// TIA Portal V20 export
// export: Created 2026-10-19T18:45:22.4932904Z, ExportSetting None, DisplayName Totally Integrated Automation Portal, DisplayVersion V20 Update 6, DisplayName TIA Portal Openness, DisplayVersion V20 Update 6, DisplayName TIA Portal Version Control Interface, DisplayVersion V20 Update 6, DisplayName SINAMICS Startdrive Advanced, DisplayVersion V20 SP1, DisplayName SINAMICS Startdrive G130, G150, S120, S150, SINAMICS MV, G220, S200, S210, DisplayVersion V20 SP1, DisplayName SINAMICS Startdrive G110M, G120, G120C, G120D, G120P, G115D, DisplayVersion V20 SP1, DisplayName STEP 7 Professional, DisplayVersion V20 Update 6, DisplayName STEP 7 Safety, DisplayVersion V20 Update 2, DisplayName WinCC Basic/Comfort/Advanced, DisplayVersion V20 Update 6, DisplayName WinCC Unified, DisplayVersion V20 Update 6
VAR_GLOBAL   // PLC tag table "IO_VFDs_1"
   VTD1_ControlWord AT %QW40 : Word;
   VTD1_StatusWord AT %IW44 : Word;
   VTD1_ActualSpeed AT %IW46 : Word;
   VTD1_ActualCurrent AT %IW48 : Word;
   VTD1_ActualTorque AT %IW50 : Word;
   VTD1_AccFactor AT %QW1513 : Word;
   C1105_Inputs AT %IW166 : Word;
   C1204_Inputs AT %IW251 : Word;
   CVTD1_Inputs AT %IW22 : Word;
   C1202_Inputs AT %IW227 : Word;
   C1103_Inputs AT %IW114 : Word;
   C1102_Inputs AT %IW38 : Word;
   C1104_Inputs AT %IW126 : Word;
   C1203_Inputs AT %IW239 : Word;
   C1206_Inputs AT %IW279 : Word;
   C1205_Inputs AT %IW263 : Word;
   C1106_Inputs AT %IW215 : Word;
   C1203_ActualTorque AT %IW235 : Word;
   C1204_ActualSpeed AT %IW243 : Word;
   C1202_StatusWord AT %IW217 : Word;
   C1206_ActualTorque AT %IW275 : Word;
   C1104_ControlWord AT %QW36 : Word;
   C1105_ActualSpeed AT %IW158 : Word;
   C1205_ControlWord AT %QW90 : Word;
   C1104_ActualCurrent AT %IW120 : Word;
   C1106_ActualSpeed AT %IW207 : Word;
   C1106_StatusWord AT %IW205 : Word;
   C1202_ControlWord AT %QW66 : Word;
   C1202_ActualSpeed AT %IW219 : Word;
   C1205_ActualCurrent AT %IW257 : Word;
   CVTD1_ActualCurrent AT %IW16 : Word;
   C1102_ActualCurrent AT %IW32 : Word;
   C1102_ActualTorque AT %IW34 : Word;
   C1205_ActualSpeed AT %IW255 : Word;
   CVTD1_ActualSpeed AT %IW14 : Word;
   C1103_ControlWord AT %QW28 : Word;
   C1106_ActualCurrent AT %IW209 : Word;
   C1204_ActualCurrent AT %IW245 : Word;
   C1105_ControlWord AT %QW50 : Word;
   C1103_ActualTorque AT %IW110 : Word;
   C1204_ControlWord AT %QW82 : Word;
   C1104_ActualSpeed AT %IW118 : Word;
   C1104_ActualTorque AT %IW122 : Word;
   C1203_ControlWord AT %QW74 : Word;
   C1204_StatusWord AT %IW241 : Word;
   C1105_ActualTorque AT %IW162 : Word;
   C1203_ActualSpeed AT %IW231 : Word;
   C1104_StatusWord AT %IW116 : Word;
   C1106_ActualTorque AT %IW211 : Word;
   C1203_StatusWord AT %IW229 : Word;
   C1202_ActualTorque AT %IW223 : Word;
   C1206_StatusWord AT %IW269 : Word;
   C1102_ControlWord AT %QW20 : Word;
   C1202_ActualCurrent AT %IW221 : Word;
   C1103_ActualSpeed AT %IW106 : Word;
   C1106_ControlWord AT %QW58 : Word;
   CVTD1_MainSetpoint AT %QW14 : Word;
   C1103_ActualCurrent AT %IW108 : Word;
   CVTD1_ActualTorque AT %IW18 : Word;
   C1105_ActualCurrent AT %IW160 : Word;
   C1105_StatusWord AT %IW156 : Word;
   CVTD1_StatusWord AT %IW12 : Word;
   C1203_ActualCurrent AT %IW233 : Word;
   C1206_ActualSpeed AT %IW271 : Word;
   CVTD1_ControlWord AT %QW12 : Word;
   C1205_ActualTorque AT %IW259 : Word;
   C1102_ActualSpeed AT %IW30 : Word;
   C1206_ControlWord AT %QW100 : Word;
   C1205_StatusWord AT %IW253 : Word;
   C1103_StatusWord AT %IW104 : Word;
   C1206_ActualCurrent AT %IW273 : Word;
   C1102_StatusWord AT %IW28 : Word;
   C1204_ActualTorque AT %IW247 : Word;
END_VAR
